# EPICS substitutions: iocs/motor/faulhaber-ioc/db/MCDC2805.substitutions
# C's iocFaulhaber MCDC2805.substitutions, P and C from st.cmd.
file "$(MOTOR)/db/motor.db"
{
pattern
{N, M,       DTYP,       S, DESC,         EGU,     DIR, VELO, VBAS, ACCL, BDST, BVEL, BACC, MRES, PREC, DHLM, DLLM, INIT}
{1, "m$(N)", "MCDC2805", 0, "motor $(N)", degrees, Pos, 10,   0.,   1.,   0,    1,    .2,   1e-3, 3,    100,  -100, ""}
}
